Fanuc KAREL source: KA00081.KL

PROGRAM KA00081
%NOLOCKGROUP
VAR
  SRC: XYZWPREXT
  DST: VECTOR
BEGIN
  SRC.X = 1.0
  DST = SRC
END KA00081
